(* PLC project OpenAI1.project, CODESYS CODESYS V3.5 SP20 *)
(* stored: creationDateTime 2026-10-15T18:40:57.5469645, modificationDateTime 2026-10-15T18:40:25.3898363 *)

PROGRAM PLC_PRG
  VAR_INPUT
    i_bStart : BOOL;
    i_bStop : BOOL;
    i_wTempSensor : INT;
  END_VAR
  VAR_OUTPUT
    o_bHeater : BOOL;
    o_bMixer : BOOL;
    o_rAvgTemp : REAL;
  END_VAR
  VAR
    a_rTempHistory : ARRAY[0..4] OF REAL;
    fbMixTimer : TON;
    i_State : INT := 0;
    i_Index : INT;
    r_Temp : REAL;
    r_Sum : REAL;
  END_VAR

                    r_Temp := (INT_TO_REAL(i_wTempSensor) * 150.0) / 27648.0;

FOR i_Index := 4 TO 1 BY -1 DO
    a_rTempHistory[i_Index] := a_rTempHistory[i_Index - 1];
END_FOR;

a_rTempHistory[0] := r_Temp;

r_Sum := 0.0;

FOR i_Index := 0 TO 4 DO
    r_Sum := r_Sum + a_rTempHistory[i_Index];
END_FOR;

o_rAvgTemp := r_Sum / 5.0;

IF NOT i_bStop THEN
    i_State := 0;
    o_bHeater := FALSE;
    o_bMixer := FALSE;
    fbMixTimer(IN := FALSE, PT := T#10s);
ELSE
    fbMixTimer(IN := (i_State = 2), PT := T#10s);

    CASE i_State OF

        0:
            o_bHeater := FALSE;
            o_bMixer := FALSE;

            IF i_bStart THEN
                i_State := 1;
            END_IF;

        1:
            o_bHeater := TRUE;
            o_bMixer := FALSE;

            IF o_rAvgTemp > 80.0 THEN
                o_bHeater := FALSE;
                o_bMixer := TRUE;
                i_State := 2;
            END_IF;

        2:
            o_bHeater := FALSE;
            o_bMixer := TRUE;

            IF fbMixTimer.Q THEN
                o_bMixer := FALSE;
                i_State := 0;
            END_IF;

        ELSE
            i_State := 0;
            o_bHeater := FALSE;
            o_bMixer := FALSE;

    END_CASE;
END_IF;
                  
END_PROGRAM

CONFIGURATION Device
  RESOURCE Application ON PLC
    TASK MainTask(INTERVAL := T#20ms, PRIORITY := 1);
    PROGRAM PLC_PRG WITH MainTask : PLC_PRG;
  END_RESOURCE
END_CONFIGURATION
